// TIA Portal V21 export
// export: Created 2026-08-21T20:18:53.8967518Z, ExportSetting None, DisplayName Totally Integrated Automation Portal, DisplayVersion V21, DisplayName STEP 7 Professional, DisplayVersion V21, DisplayName STEP 7 Safety, DisplayVersion V21, DisplayName Tech WebApplication, DisplayVersion V21, DisplayName WinCC Basic/Comfort/Advanced, DisplayVersion V21, DisplayName WinCC Professional, DisplayVersion V21, DisplayName WinCC Unified, DisplayVersion V21
FUNCTION_BLOCK "MTPAnaMon_Type1"   // FB15, FBD
{ S7_Optimized_Access := 'TRUE' }
// stored: MemoryReserve 100, SetENOAutomatically false
   VAR_INPUT
      PV { ExternalAccessible := 'False'; ExternalVisible := 'False'; ExternalWritable := 'False'} : Word;
      PV_QB { ExternalAccessible := 'False'; ExternalVisible := 'False'; ExternalWritable := 'False'} : Bool := true;
      PV_Unit { ExternalAccessible := 'False'; ExternalVisible := 'False'; ExternalWritable := 'False'} : Int := 1001;
      PV_AH_En { ExternalAccessible := 'False'; ExternalVisible := 'False'; ExternalWritable := 'False'} : Bool := true;
      PV_WH_En { ExternalAccessible := 'False'; ExternalVisible := 'False'; ExternalWritable := 'False'} : Bool := true;
      PV_TH_En { ExternalAccessible := 'False'; ExternalVisible := 'False'; ExternalWritable := 'False'} : Bool;
      PV_TL_En { ExternalAccessible := 'False'; ExternalVisible := 'False'; ExternalWritable := 'False'} : Bool;
      PV_WL_En { ExternalAccessible := 'False'; ExternalVisible := 'False'; ExternalWritable := 'False'} : Bool := true;
      PV_AL_En { ExternalAccessible := 'False'; ExternalVisible := 'False'; ExternalWritable := 'False'} : Bool := true;
   END_VAR
   VAR_OUTPUT
      to_Indicate { ExternalAccessible := 'False'; ExternalVisible := 'False'; ExternalWritable := 'False'} : "StruCm";
   END_VAR
   VAR
      AnIn_IDB { ExternalAccessible := 'False'; ExternalVisible := 'False'; ExternalWritable := 'False'} : "AnIn";
      MonAnL_IDB : "MonAnL";
      MTPAnaMon_IDB { ExternalVisible := 'False'; S7_SetPoint := 'True'} : "MTPAnaMon";
   END_VAR
   VAR_TEMP
      PV_Out : "AnaVal";
      CSF_NOP : "DigVal";
      BadAnIn : "DigVal";
      BadOut : "DigVal";
      ScaleOut : "ScaVal";
   END_VAR
   VAR_TEMP   // added for the SCL form of the ladder/FBD networks
      _w1 : Bool;
   END_VAR
BEGIN

REGION Network 1: Convert / Init
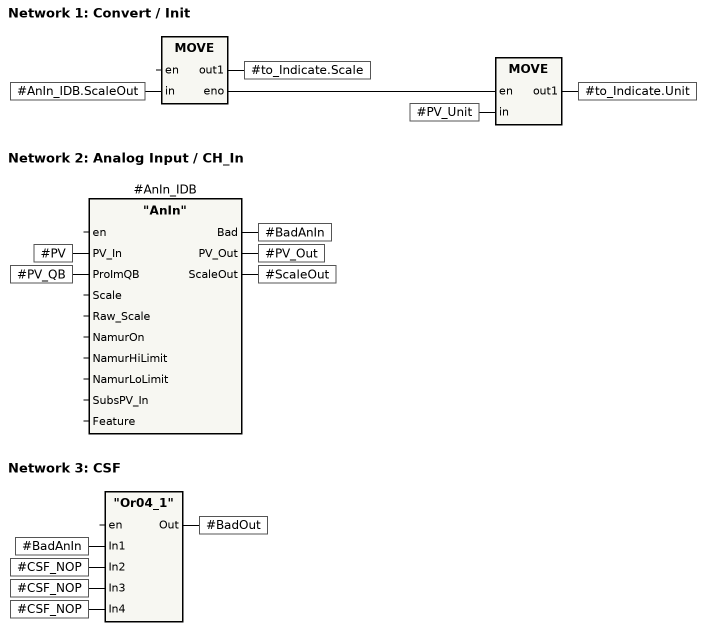
   #to_Indicate.Scale := #AnIn_IDB.ScaleOut;
   #to_Indicate.Unit := #PV_Unit;
END_REGION

REGION Network 2: Analog Input / CH_In
   #AnIn_IDB(PV_In := #PV, ProImQB := #PV_QB, Bad => #BadAnIn, PV_Out => #PV_Out, ScaleOut => #ScaleOut);   // "AnIn"
END_REGION

REGION Network 3: CSF
   "Or04_1"(In1 := #BadAnIn, In2 := #CSF_NOP, In3 := #CSF_NOP, In4 := #CSF_NOP, Out => #BadOut);
END_REGION

REGION Network 4: MonAnL
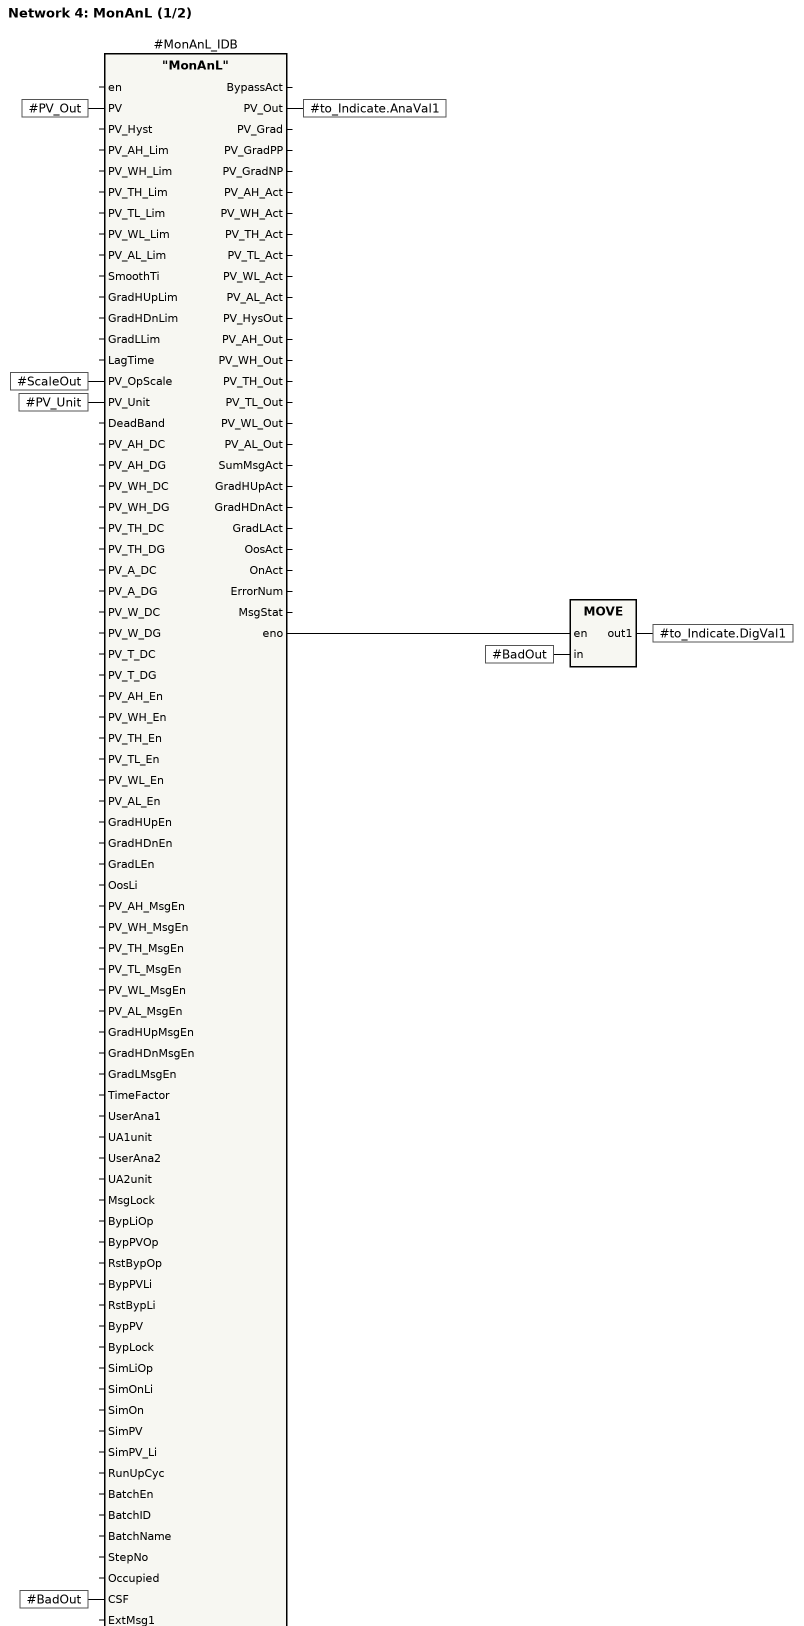
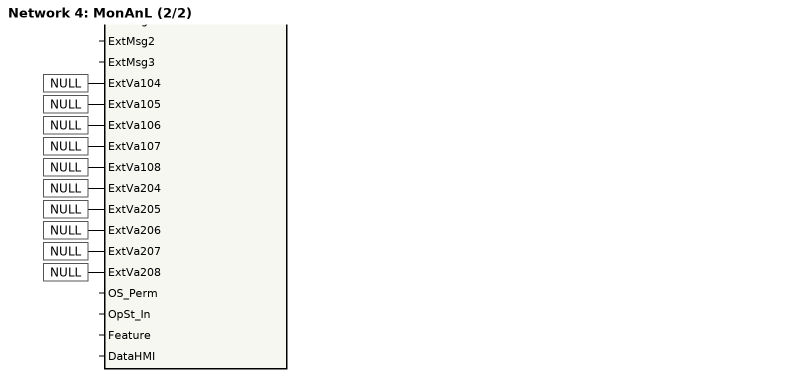
   #MonAnL_IDB(PV := #PV_Out,   // "MonAnL"
               PV_OpScale := #ScaleOut,
               PV_Unit := #PV_Unit,
               CSF := #BadOut,
               ExtVa104 := NULL,
               ExtVa105 := NULL,
               ExtVa106 := NULL,
               ExtVa107 := NULL,
               ExtVa108 := NULL,
               ExtVa204 := NULL,
               ExtVa205 := NULL,
               ExtVa206 := NULL,
               ExtVa207 := NULL,
               ExtVa208 := NULL,
               PV_Out => #to_Indicate.AnaVal1,
               ENO => #_w1);
   IF #_w1 THEN #to_Indicate.DigVal1 := #BadOut; END_IF;
END_REGION

REGION Network 5: MTP / MTP Connector block
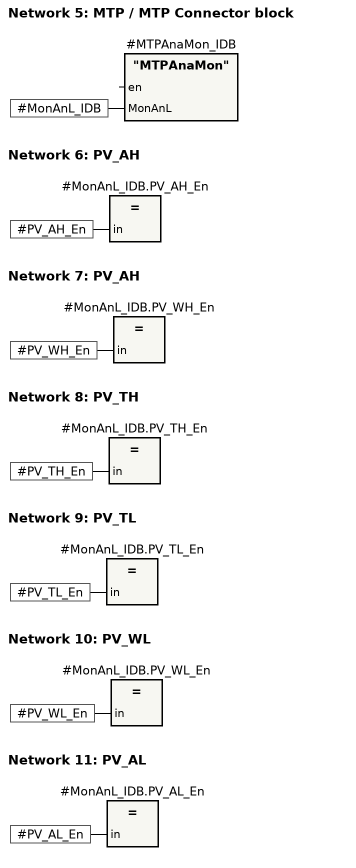
   #MTPAnaMon_IDB(MonAnL := #MonAnL_IDB);   // "MTPAnaMon"
END_REGION

REGION Network 6: PV_AH
   #MonAnL_IDB.PV_AH_En := #PV_AH_En;
END_REGION

REGION Network 7: PV_AH
   #MonAnL_IDB.PV_WH_En := #PV_WH_En;
END_REGION

REGION Network 8: PV_TH
   #MonAnL_IDB.PV_TH_En := #PV_TH_En;
END_REGION

REGION Network 9: PV_TL
   #MonAnL_IDB.PV_TL_En := #PV_TL_En;
END_REGION

REGION Network 10: PV_WL
   #MonAnL_IDB.PV_WL_En := #PV_WL_En;
END_REGION

REGION Network 11: PV_AL
   #MonAnL_IDB.PV_AL_En := #PV_AL_En;
END_REGION
END_FUNCTION_BLOCK
